(* IEC 61131-3 sources: codesys-ai-industrial-robot-control/plc/src/Framework/FB_PartQueue, 6 files *)

(* ---- AddRecord.st ---- *)
// Stores the record in a free slot. Returns its index, or 0 when the queue is full.
METHOD AddRecord : UINT
VAR_INPUT
    stRec : ST_PartRecord;
END_VAR
VAR
    i : UINT;
END_VAR

AddRecord := 0;
FOR i := 1 TO GVL_Config.MAX_PARTS DO
    IF aRecords[i].eState = E_PartState.Free THEN
        aRecords[i] := stRec;
        AddRecord := i;
        RETURN;
    END_IF
END_FOR

(* ---- Clear.st ---- *)
// Empty every slot.
METHOD Clear
VAR
    i : UINT;
END_VAR

FOR i := 1 TO GVL_Config.MAX_PARTS DO
    aRecords[i] := stEmpty;
END_FOR

(* ---- FindIndex.st ---- *)
// Index of the record with this part id, or 0.
METHOD FindIndex : UINT
VAR_INPUT
    udiPartId : UDINT;
END_VAR
VAR
    i : UINT;
END_VAR

FindIndex := 0;
IF udiPartId = 0 THEN
    RETURN;
END_IF
FOR i := 1 TO GVL_Config.MAX_PARTS DO
    IF aRecords[i].eState <> E_PartState.Free AND aRecords[i].udiPartId = udiPartId THEN
        FindIndex := i;
        RETURN;
    END_IF
END_FOR

(* ---- GetRecord.st ---- *)
METHOD GetRecord : ST_PartRecord
VAR_INPUT
    uiIdx : UINT;
END_VAR

IF uiIdx >= 1 AND uiIdx <= GVL_Config.MAX_PARTS THEN
    GetRecord := aRecords[uiIdx];
ELSE
    GetRecord := stEmpty;
END_IF

(* ---- PutRecord.st ---- *)
METHOD PutRecord
VAR_INPUT
    uiIdx : UINT;
    stRec : ST_PartRecord;
END_VAR

IF uiIdx >= 1 AND uiIdx <= GVL_Config.MAX_PARTS THEN
    aRecords[uiIdx] := stRec;
END_IF

(* ---- Release.st ---- *)
METHOD Release
VAR_INPUT
    uiIdx : UINT;
END_VAR

IF uiIdx >= 1 AND uiIdx <= GVL_Config.MAX_PARTS THEN
    aRecords[uiIdx] := stEmpty;
END_IF
